(* IEC 61131-3 sources: plcassist-cli/packages/volt-lsp-iec/test-corpus/lenze-mid/Device/Plc Logic/Application/Library Manager/StringUtils, 60 files *)

(* ---- CONSTANTS.gvl ---- *)
VAR_GLOBAL
	NULL : POINTER TO BYTE := 0;
END_VAR

(* ---- GVL_UTF8.gvl ---- *)
VAR_GLOBAL
	TRAILINGBYTESFORUTF8 : ARRAY [0..255] OF BYTE := [0, 0, 0, 0, 0, 0, 0, 0, 0, 0, 0, 0, 0, 0, 0, 0, 0, 0, 0, 0, 0, 0, 0, 0, 0, 0, 0, 0, 0, 0, 0, 0, 0, 0, 0, 0, 0, 0, 0, 0, 0, 0, 0, 0, 0, 0, 0, 0, 0, 0, 0, 0, 0, 0, 0, 0, 0, 0, 0, 0, 0, 0, 0, 0, 0, 0, 0, 0, 0, 0, 0, 0, 0, 0, 0, 0, 0, 0, 0, 0, 0, 0, 0, 0, 0, 0, 0, 0, 0, 0, 0, 0, 0, 0, 0, 0, 0, 0, 0, 0, 0, 0, 0, 0, 0, 0, 0, 0, 0, 0, 0, 0, 0, 0, 0, 0, 0, 0, 0, 0, 0, 0, 0, 0, 0, 0, 0, 0, 0, 0, 0, 0, 0, 0, 0, 0, 0, 0, 0, 0, 0, 0, 0, 0, 0, 0, 0, 0, 0, 0, 0, 0, 0, 0, 0, 0, 0, 0, 0, 0, 0, 0, 0, 0, 0, 0, 0, 0, 0, 0, 0, 0, 0, 0, 0, 0, 0, 0, 0, 0, 0, 0, 0, 0, 0, 0, 0, 0, 0, 0, 0, 0, 1, 1, 1, 1, 1, 1, 1, 1, 1, 1, 1, 1, 1, 1, 1, 1, 1, 1, 1, 1, 1, 1, 1, 1, 1, 1, 1, 1, 1, 1, 1, 1, 2, 2, 2, 2, 2, 2, 2, 2, 2, 2, 2, 2, 2, 2, 2, 2, 3, 3, 3, 3, 3, 3, 3, 3, 4, 4, 4, 4, 5, 5, 5, 5];
	FIRSTBYTEMARK : ARRAY [0..6] OF BYTE := [16#0, 16#0, 16#C0, 16#E0, 16#F0, 16#F8, 16#FC];
	OFFSETSFROMUTF8 : ARRAY [0..5] OF DWORD := [16#0, 16#3080, 16#E2080, 16#3C82080, 16#FA082080, 16#82082080];
	HALFSHIFT : INT := 10;
	HALFBASE : DWORD := 16#10000;
	HALFMASK : DWORD := 16#3FF;
	UNI_REPLACEMENT_CHAR : DWORD := 16#FFFD;
	UNI_MAX_BMP : DWORD := 16#FFFF;
	UNI_MAX_UTF16 : DWORD := 16#10FFFF;
	UNI_MAX_UTF32 : DWORD := 16#7FFFFFFF;
	UNI_MAX_LEGAL_UTF32 : DWORD := 16#10FFFF;
	BYTEMASK : DWORD := 16#BF;
	BYTEMARK : DWORD := 16#80;
	UNI_SUR_HIGH_START : DWORD := 16#D800;
	UNI_SUR_HIGH_END : DWORD := 16#DBFF;
	UNI_SUR_LOW_START : DWORD := 16#DC00;
	UNI_SUR_LOW_END : DWORD := 16#DFFF;
	ERR_SOURCE_EXHAUSTED : UDINT := 16#40A0;
	ERR_TARGET_EXHAUSTED : UDINT := 16#40A1;
	ERR_SOURCE_ILLEGAL : UDINT := 16#40A2;
END_VAR

(* ---- PLACEHOLDERCONSTANTS.gvl ---- *)
VAR_GLOBAL
	DFMT_FIRST_PLACEHOLDER : EDateTimePlaceholder := EDateTimePlaceholder.DFMT_5_DIGIT_DAY;
	DFMT_LAST_PLACEHOLDER : EDateTimePlaceholder := EDateTimePlaceholder.DFMT_1_DIGIT_YEAR;
	TFMT_FIRST_PLACEHOLDER : EDateTimePlaceholder := EDateTimePlaceholder.TFMT_2_DIGIT_HOUR_24_HOUR_CLOCK;
	TFMT_LAST_PLACEHOLDER : EDateTimePlaceholder := EDateTimePlaceholder.TFMT_1_DIGIT_ZONE_DESIGNATOR;
END_VAR

(* ---- STRINGUTILSVERSIONCONSTANTS.gvl ---- *)
VAR_GLOBAL
	_STRINGUTILS_VERSION_LARGEROREQUAL_3_5_3_40_ : INT := 0;
END_VAR

(* ---- ICHARBUFFERSTRING.itf ---- *)
INTERFACE ICHARBUFFERSTRING
END_INTERFACE

METHOD ASWSTRING : CharBufferPtr
END_METHOD

METHOD COPY : DINT
VAR_INPUT
	CBSSOURCE : REFERENCE TO CharBufferString;
END_VAR
END_METHOD

METHOD FROMSTRING : BOOL
VAR_INPUT
	STSTRING : STRING(255);
END_VAR
END_METHOD

METHOD INITCONVERTED : BOOL
VAR_INPUT
	PBUFFER : POINTER TO BYTE;
	UIBUFFERSIZE : UINT;
END_VAR
END_METHOD

(* ---- ILOCALIZEDDATETIMENAMES.itf ---- *)
INTERFACE ILOCALIZEDDATETIMENAMES
END_INTERFACE

METHOD GETDAYLONG : CharBufferPtr
VAR_INPUT
	UIDAYOFWEEK : UINT;
END_VAR
END_METHOD

METHOD GETDAYSHORT : CharBufferPtr
VAR_INPUT
	UIDAYOFWEEK : UINT;
END_VAR
END_METHOD

METHOD GETMONTHLONG : CharBufferPtr
VAR_INPUT
	UIMONTH : UINT;
END_VAR
END_METHOD

METHOD GETMONTHSHORT : CharBufferPtr
VAR_INPUT
	UIMONTH : UINT;
END_VAR
END_METHOD

(* ---- _PRINTF.fun ---- *)
FUNCTION _PRINTF : BOOL
VAR_INPUT
	CBPRESULT : CharBufferPtr;
	UIRESULTCAPACITY : UINT;
	STRINGTYPE : __SYSTEM.TYPE_CLASS;
	CBPFORMAT : CharBufferPtr;
	PVALUE : POINTER TO BYTE;
	TYPECLASS : __SYSTEM.TYPE_CLASS;
END_VAR
END_FUNCTION

(* ---- ANALYZEPLACEHOLDERS.fun ---- *)
FUNCTION ANALYZEPLACEHOLDERS : EPlaceholderAnalyzationState
VAR_INPUT
	RCBSMESSAGE : REFERENCE TO CharBufferString;
	PAPLACEHOLDERS : POINTER TO ARRAY [0..0] OF PlaceholderDescription;
	ICOUNTPLACEHOLDERTOCHECK : INT;
	PAPLACEHOLDEROCCURRENCE : POINTER TO ARRAY [0..0] OF DateTimePlaceholderOccurrence;
	SIMAXCOUNTPLACEHOLDERS : SINT;
END_VAR
VAR_OUTPUT
	SICOUNTPLACEHOLDERS : SINT;
END_VAR
END_FUNCTION

(* ---- ANALYZEPLACEHOLDERSDATETIME.fun ---- *)
FUNCTION ANALYZEPLACEHOLDERSDATETIME : EPlaceholderAnalyzationState
VAR_INPUT
	RCBSMESSAGE : REFERENCE TO CharBufferString;
	PAPLACEHOLDERS : POINTER TO ARRAY [0..0] OF PlaceholderDescription;
	ICOUNTPLACEHOLDERTOCHECK : INT;
	PAPLACEHOLDEROCCURRENCE : POINTER TO ARRAY [0..0] OF DateTimePlaceholderOccurrence;
	SIMAXCOUNTPLACEHOLDERS : SINT;
END_VAR
VAR_OUTPUT
	SICOUNTPLACEHOLDERS : SINT;
END_VAR
END_FUNCTION

(* ---- CHARACTERATEQUALS.fun ---- *)
FUNCTION CHARACTERATEQUALS : BOOL
VAR_INPUT
	CBSSOURCE : REFERENCE TO CharBufferString;
	IPOSITION : INT;
	STCHAR : STRING(1);
END_VAR
END_FUNCTION

(* ---- CHARTOUPPER.fun ---- *)
FUNCTION CHARTOUPPER : BYTE
VAR_INPUT
	BYCHAR : BYTE;
END_VAR
END_FUNCTION

(* ---- CONVERTUTF16TOUTF8.fun ---- *)
FUNCTION CONVERTUTF16TOUTF8 : UDINT
VAR_INPUT
	SOURCESTART : POINTER TO WORD;
	TARGETSTART : POINTER TO BYTE;
	DWTARGETBUFFERSIZE : DWORD;
	BSTRICTCONVERSION : BOOL;
END_VAR
END_FUNCTION

(* ---- CONVERTUTF8TOUTF16.fun ---- *)
FUNCTION CONVERTUTF8TOUTF16 : UDINT
VAR_INPUT
	SOURCESTART : POINTER TO BYTE;
	TARGETSTART : POINTER TO WORD;
	DWTARGETBUFFERSIZE : DWORD;
	BSTRICTCONVERSION : BOOL;
END_VAR
END_FUNCTION

(* ---- HELPISSAMEIGNORECASE.fun ---- *)
FUNCTION HELPISSAMEIGNORECASE : BOOL
VAR_INPUT
	BY1 : BYTE;
	BY2 : BYTE;
END_VAR
END_FUNCTION

(* ---- HELPSTRCMPENDA.fun ---- *)
FUNCTION HELPSTRCMPENDA : BOOL
VAR_INPUT
	PCOMPLETETEXT : CharBufferPtr;
	PSUBTEXT : CharBufferPtr;
	XIGNORECASE : BOOL;
END_VAR
END_FUNCTION

(* ---- HELPSTRCMPSTARTA.fun ---- *)
FUNCTION HELPSTRCMPSTARTA : BOOL
VAR_INPUT
	PCOMPLETETEXT : CharBufferPtr;
	PSUBTEXT : CharBufferPtr;
	XIGNORECASE : BOOL;
END_VAR
END_FUNCTION

(* ---- HELPTRIM.fun ---- *)
FUNCTION HELPTRIM : POINTER TO BYTE
VAR_INPUT
	PTEXT : CharBufferPtr;
	XTRIMLEFT : BOOL;
END_VAR
END_FUNCTION

(* ---- HELPTRIMW.fun ---- *)
FUNCTION HELPTRIMW : POINTER TO WORD
VAR_INPUT
	PTEXT : CharBufferPtr;
	XTRIMLEFT : BOOL;
END_VAR
END_FUNCTION

(* ---- ISLEGALUTF8.fun ---- *)
FUNCTION ISLEGALUTF8 : BOOL
VAR_INPUT
	SOURCE : POINTER TO BYTE;
	LENGTH : INT;
END_VAR
END_FUNCTION

(* ---- ISSPACECHARACTER.fun ---- *)
FUNCTION ISSPACECHARACTER : BOOL
VAR_INPUT
	WCHARACTER : WORD;
END_VAR
END_FUNCTION

(* ---- STRCASECMPA.fun ---- *)
FUNCTION STRCASECMPA : INT
VAR_INPUT
	PBYTE1 : POINTER TO BYTE;
	PBYTE2 : POINTER TO BYTE;
END_VAR
END_FUNCTION

(* ---- STRCASECMPENDA.fun ---- *)
FUNCTION STRCASECMPENDA : INT
VAR_INPUT
	PSTRING : CharBufferPtr;
	PSUFFIX : CharBufferPtr;
END_VAR
END_FUNCTION

(* ---- STRCASECMPSTARTA.fun ---- *)
FUNCTION STRCASECMPSTARTA : INT
VAR_INPUT
	PSTRING : CharBufferPtr;
	PPREFIX : CharBufferPtr;
END_VAR
END_FUNCTION

(* ---- STRCASECMPW.fun ---- *)
FUNCTION STRCASECMPW : INT
VAR_INPUT
	PWD1 : POINTER TO WORD;
	PWD2 : POINTER TO WORD;
END_VAR
END_FUNCTION

(* ---- STRCASEFINDA.fun ---- *)
FUNCTION STRCASEFINDA : INT
VAR_INPUT
	PST1 : POINTER TO STRING(255);
	PST2 : POINTER TO STRING(255);
	UISEARCHSTART : UINT;
END_VAR
END_FUNCTION

(* ---- STRCASEFINDW.fun ---- *)
FUNCTION STRCASEFINDW : INT
VAR_INPUT
	PST1 : POINTER TO WSTRING(255);
	PST2 : POINTER TO WSTRING(255);
	UISEARCHSTART : UINT;
END_VAR
END_FUNCTION

(* ---- STRCMP.fun ---- *)
FUNCTION STRCMP : DINT
VAR_INPUT
	CBSSTRING1 : REFERENCE TO CharBufferString;
	CBSSTRING2 : REFERENCE TO CharBufferString;
END_VAR
END_FUNCTION

(* ---- STRCMPA.fun ---- *)
FUNCTION STRCMPA : INT
VAR_INPUT
	PBY1 : POINTER TO BYTE;
	PBY2 : POINTER TO BYTE;
END_VAR
END_FUNCTION

(* ---- STRCMPENDA.fun ---- *)
FUNCTION STRCMPENDA : INT
VAR_INPUT
	PSTRING : CharBufferPtr;
	PSUFFIX : CharBufferPtr;
END_VAR
END_FUNCTION

(* ---- STRCMPSTARTA.fun ---- *)
FUNCTION STRCMPSTARTA : INT
VAR_INPUT
	PSTRING : CharBufferPtr;
	PPREFIX : CharBufferPtr;
END_VAR
END_FUNCTION

(* ---- STRCMPW.fun ---- *)
FUNCTION STRCMPW : INT
VAR_INPUT
	PWD1 : POINTER TO WORD;
	PWD2 : POINTER TO WORD;
END_VAR
END_FUNCTION

(* ---- STRCONCATA.fun ---- *)
FUNCTION STRCONCATA : BOOL
VAR_INPUT
	PSTFROM : CharBufferPtr;
	PSTTO : CharBufferPtr;
	IBUFFERSIZE : INT;
END_VAR
END_FUNCTION

(* ---- STRCONCATW.fun ---- *)
FUNCTION STRCONCATW : BOOL
VAR_INPUT
	PSTFROM : CharBufferPtr;
	PSTTO : CharBufferPtr;
	IBUFFERSIZE : INT;
END_VAR
END_FUNCTION

(* ---- STRCPY.fun ---- *)
FUNCTION STRCPY : DINT
VAR_INPUT
	CBSTARGET : REFERENCE TO CharBufferString;
	CBSSOURCE : REFERENCE TO CharBufferString;
END_VAR
END_FUNCTION

(* ---- STRCPYA.fun ---- *)
FUNCTION STRCPYA : DINT
VAR_INPUT
	PBUFFER : CharBufferPtr;
	IBUFFERSIZE : DINT;
	PSTR : CharBufferPtr;
END_VAR
END_FUNCTION

(* ---- STRCPYFROM.fun ---- *)
FUNCTION STRCPYFROM : DINT
VAR_INPUT
	RCBSTARGET : REFERENCE TO CharBufferString;
	RCBSSOURCE : REFERENCE TO CharBufferString;
	DISOURCEOFFSET : DINT;
	DITARGETOFFSET : DINT;
	DICOUNTCHARACTERS : DINT;
END_VAR
END_FUNCTION

(* ---- STRCPYW.fun ---- *)
FUNCTION STRCPYW : DINT
VAR_INPUT
	PBUFFER : CharBufferPtr;
	IBUFFERSIZE : DINT;
	PSTR : CharBufferPtr;
END_VAR
END_FUNCTION

(* ---- STRFIND.fun ---- *)
FUNCTION STRFIND : INT
VAR_INPUT
	CBSSOURCE : REFERENCE TO CharBufferString;
	CBSTOSEARCHFOR : REFERENCE TO CharBufferString;
END_VAR
END_FUNCTION

(* ---- STRFINDA.fun ---- *)
FUNCTION STRFINDA : INT
VAR_INPUT
	PST1 : POINTER TO STRING(255);
	PST2 : POINTER TO STRING(255);
	UISEARCHSTART : UINT;
END_VAR
END_FUNCTION

(* ---- STRFINDFROM.fun ---- *)
FUNCTION STRFINDFROM : INT
VAR_INPUT
	CBSSOURCE : REFERENCE TO CharBufferString;
	CBSTOSEARCHFOR : REFERENCE TO CharBufferString;
	ISEARCHSTART : UINT;
END_VAR
END_FUNCTION

(* ---- STRFINDW.fun ---- *)
FUNCTION STRFINDW : INT
VAR_INPUT
	PST1 : POINTER TO WSTRING(255);
	PST2 : POINTER TO WSTRING(255);
	UISEARCHSTART : UINT;
END_VAR
END_FUNCTION

(* ---- STRINGTOCHARBUFFERPTR.fun ---- *)
FUNCTION STRINGTOCHARBUFFERPTR : BOOL
VAR_INPUT
	STSTRING : STRING(255);
	CBSRESULT : REFERENCE TO CharBufferString;
END_VAR
END_FUNCTION

(* ---- STRISNULLOREMPTYA.fun ---- *)
FUNCTION STRISNULLOREMPTYA : BOOL
VAR_INPUT
	PSTDATA : CharBufferPtr;
END_VAR
END_FUNCTION

(* ---- STRISNULLOREMPTYW.fun ---- *)
FUNCTION STRISNULLOREMPTYW : BOOL
VAR_INPUT
	PSTDATA : CharBufferPtr;
END_VAR
END_FUNCTION

(* ---- STRLEN.fun ---- *)
FUNCTION STRLEN : DINT
VAR_INPUT
	CBSSOURCE : REFERENCE TO CharBufferString;
END_VAR
END_FUNCTION

(* ---- STRLENA.fun ---- *)
FUNCTION STRLENA : DINT
VAR_INPUT
	PSTDATA : CharBufferPtr;
END_VAR
END_FUNCTION

(* ---- STRLENW.fun ---- *)
FUNCTION STRLENW : DINT
VAR_INPUT
	PSTDATA : CharBufferPtr;
END_VAR
END_FUNCTION

(* ---- STRPADLEFTA.fun ---- *)
FUNCTION STRPADLEFTA : BOOL
VAR_INPUT
	BYPADCHAR : BYTE;
	PSTFROM : CharBufferPtr;
	PSTTO : CharBufferPtr;
	DIBUFFERSIZE : DINT;
END_VAR
END_FUNCTION

(* ---- STRPADLEFTW.fun ---- *)
FUNCTION STRPADLEFTW : BOOL
VAR_INPUT
	WPADCHAR : WORD;
	PSTFROM : CharBufferPtr;
	PSTTO : CharBufferPtr;
	DIBUFFERSIZE : DINT;
END_VAR
END_FUNCTION

(* ---- STRPADRIGHTA.fun ---- *)
FUNCTION STRPADRIGHTA : BOOL
VAR_INPUT
	BYPADCHAR : BYTE;
	PSTFROM : CharBufferPtr;
	PSTTO : CharBufferPtr;
	DIBUFFERSIZE : DINT;
END_VAR
END_FUNCTION

(* ---- STRPADRIGHTW.fun ---- *)
FUNCTION STRPADRIGHTW : BOOL
VAR_INPUT
	WPADCHAR : WORD;
	PSTFROM : CharBufferPtr;
	PSTTO : CharBufferPtr;
	DIBUFFERSIZE : DINT;
END_VAR
END_FUNCTION

(* ---- STRTRIMW.fun ---- *)
FUNCTION STRTRIMW : BOOL
VAR_INPUT
	PSTRING : CharBufferPtr;
END_VAR
END_FUNCTION

(* ---- STUSPRINTF.fun ---- *)
FUNCTION STUSPRINTF : INT
VAR_INPUT
	PSTFORMAT : POINTER TO STRING;
	PVARADR : POINTER TO DWORD;
	UDIVARTYPE : __SYSTEM.TYPE_CLASS;
	PBUFFER : POINTER TO BYTE;
	DWBUFFERSIZE : UDINT;
END_VAR
END_FUNCTION

(* ---- STUSPRINTFW.fun ---- *)
FUNCTION STUSPRINTFW : INT
VAR_INPUT
	WSTFORMAT : POINTER TO WSTRING;
	PVARADR : POINTER TO DWORD;
	UDIVARTYPE : __SYSTEM.TYPE_CLASS;
	PBUFFER : POINTER TO BYTE;
	DWBUFFERSIZE : UDINT;
END_VAR
END_FUNCTION

(* ---- WCHARTOUPPER.fun ---- *)
FUNCTION WCHARTOUPPER : WORD
VAR_INPUT
	WDCHAR : WORD;
END_VAR
END_FUNCTION

(* ---- ABSTRACTFORMATTER.fb ---- *)
FUNCTION_BLOCK ABSTRACTFORMATTER
VAR
	M_APLACEHOLDEROCCURRENCE : ARRAY [0..(COUNT_PLACEHOLDERS_IN_FORMAT_STRING - 1)] OF DateTimePlaceholderOccurrence;
	M_SICOUNTPLACEHOLDERS : SINT := -1;
	M_EPLACEHOLDERANALYZATIONSTATE : EPlaceholderAnalyzationState;
	M_SFORMATSTRING : STRING(50);
	M_IFORMATSTRINGLENGTH : INT;
	COUNT_PLACEHOLDERS_IN_FORMAT_STRING : INT := 10;
	COUNT_PLACEHOLDERS_IN_DATETIMEFORMAT_STRING : INT := 20;
	MAX_FORMAT_STRING_LENGTH : SINT := 50;
END_VAR
END_FUNCTION_BLOCK

(* ---- CHARBUFFERSTRING.fb ---- *)
FUNCTION_BLOCK CHARBUFFERSTRING
VAR_INPUT
	M_UIBUFFERSIZE : UINT;
	M_CBPBUFFER : CharBufferPtr;
	M_TYPE : __SYSTEM.TYPE_CLASS;
	M_ASSTRING : POINTER TO STRING(255);
	M_ASWSTRING : POINTER TO WSTRING(255);
	M_BALLOCATED : BOOL;
END_VAR
VAR
	CAPACITY : UINT;
	CHARACTERS : CharBufferPtr;
	LENGTH : DINT;
	STRINGTYPE : __SYSTEM.TYPE_CLASS;
END_VAR
END_FUNCTION_BLOCK

METHOD ASWSTRING : CharBufferPtr
END_METHOD

METHOD CHARAT : BYTE
VAR_INPUT
	IPOSITION : INT;
END_VAR
END_METHOD

METHOD CHARATEQUALS : BOOL
VAR_INPUT
	IPOSITION : INT;
	STCHAR : STRING(1);
END_VAR
END_METHOD

METHOD COPY : DINT
VAR_INPUT
	CBSSOURCE : REFERENCE TO CharBufferString;
END_VAR
END_METHOD

METHOD COPYFROM
VAR_INPUT
	RCBSSOURCE : REFERENCE TO CharBufferString;
	DISOURCEOFFSET : DINT;
	DITARGETOFFSET : DINT;
	DICOUNTCHARACTERS : DINT;
END_VAR
END_METHOD

METHOD COPYFROM2 : DINT
VAR_INPUT
	RSSOURCE : REFERENCE TO STRING(255);
	DITARGETOFFSET : DINT;
END_VAR
END_METHOD

METHOD DELETE : DINT
VAR_INPUT
	ILENGTH : INT;
	IPOSITION : INT;
END_VAR
END_METHOD

METHOD FB_EXIT : BOOL
VAR_INPUT
	BINCOPYCODE : BOOL;
END_VAR
END_METHOD

METHOD FB_INIT : BOOL
VAR_INPUT
	BINITRETAINS : BOOL;
	BINCOPYCODE : BOOL;
	UIBUFFERSIZE : UINT;
	STRINGTYPE : __SYSTEM.TYPE_CLASS;
END_VAR
END_METHOD

METHOD FIND : INT
VAR_INPUT
	CBSTOSEARCHFOR : REFERENCE TO CharBufferString;
END_VAR
END_METHOD

METHOD FINDFROM : INT
VAR_INPUT
	CBSTOSEARCHFOR : REFERENCE TO CharBufferString;
	ISEARCHSTART : UINT;
END_VAR
END_METHOD

METHOD FROMSTRING : BOOL
VAR_INPUT
	STSTRING : STRING(255);
END_VAR
END_METHOD

METHOD INIT : BOOL
VAR_INPUT
	PBUFFER : POINTER TO BYTE;
	UIBUFFERSIZE : UINT;
	STRINGTYPE : __SYSTEM.TYPE_CLASS;
END_VAR
END_METHOD

METHOD INITCONVERTED : BOOL
VAR_INPUT
	PBUFFER : POINTER TO BYTE;
	UIBUFFERSIZE : UINT;
END_VAR
END_METHOD

METHOD INITIALIZE : BOOL
VAR_INPUT
	CBPSOURCE : CharBufferPtr;
	STRINGTYPE : __SYSTEM.TYPE_CLASS;
END_VAR
END_METHOD

METHOD INSERT
VAR_INPUT
	CBSINSERT : REFERENCE TO CharBufferString;
	IPOSITION : INT;
END_VAR
END_METHOD

METHOD MID
VAR_INPUT
	ILENGTH : INT;
	IPOSITION : INT;
	CBSRESULT : REFERENCE TO CharBufferString;
END_VAR
END_METHOD

METHOD PLACEHOLDEREQUALS : BOOL
VAR_INPUT
	STVALUE : STRING;
	WSTVALUE : WSTRING;
END_VAR
END_METHOD

METHOD REPLACE
VAR_INPUT
	CBSREPLACEWITH : REFERENCE TO CharBufferString;
	ILENGTHTOREPLACE : INT;
	IPOSITION : INT;
END_VAR
END_METHOD

(* ---- DATEFORMATTER.fb ---- *)
FUNCTION_BLOCK DATEFORMATTER EXTENDS AbstractFormatter
VAR
	M_CBSPLACEHOLDER2DIGITDAY : CharBufferString;
	M_CBSPLACEHOLDER1DIGITDAY : CharBufferString;
	M_CBSPLACEHOLDER2DIGITMONTH : CharBufferString;
	M_CBSPLACEHOLDER1DIGITMONTH : CharBufferString;
	M_CBSPLACEHOLDER4DIGITYEAR : CharBufferString;
	M_CBSPLACEHOLDER2DIGITYEAR : CharBufferString;
	M_CBSPLACEHOLDER1DIGITYEAR : CharBufferString;
END_VAR
END_FUNCTION_BLOCK

METHOD FB_EXIT : BOOL
VAR_INPUT
	BINCOPYCODE : BOOL;
END_VAR
END_METHOD

METHOD FB_INIT : BOOL
VAR_INPUT
	BINITRETAINS : BOOL;
	BINCOPYCODE : BOOL;
END_VAR
END_METHOD

METHOD FORMAT : STRING
VAR_INPUT
	PDATE : SYSTIMEDATE;
END_VAR
END_METHOD

METHOD SETFORMATSTRING
VAR_INPUT
	SFORMATSTRING : STRING(MAX_FORMAT_STRING_LENGTH);
END_VAR
END_METHOD

(* ---- DATETIMEFORMATTER.fb ---- *)
FUNCTION_BLOCK DATETIMEFORMATTER EXTENDS AbstractFormatter
VAR
	M_APLACEHOLDEROCCURRENCEDATETIME : ARRAY [0..(COUNT_PLACEHOLDERS_IN_DATETIMEFORMAT_STRING - 1)] OF DateTimePlaceholderOccurrence;
	M_CBSPLACEHOLDER5DIGITDAY : CharBufferString;
	M_CBSPLACEHOLDER4DIGITDAY : CharBufferString;
	M_CBSPLACEHOLDER3DIGITDAY : CharBufferString;
	M_CBSPLACEHOLDER2DIGITDAY : CharBufferString;
	M_CBSPLACEHOLDER1DIGITDAY : CharBufferString;
	M_CBSPLACEHOLDER3DIGITDAYOFYEAR : CharBufferString;
	M_CBSPLACEHOLDER4DIGITMONTH : CharBufferString;
	M_CBSPLACEHOLDER3DIGITMONTH : CharBufferString;
	M_CBSPLACEHOLDER2DIGITMONTH : CharBufferString;
	M_CBSPLACEHOLDER1DIGITMONTH : CharBufferString;
	M_CBSPLACEHOLDER4DIGITYEAR : CharBufferString;
	M_CBSPLACEHOLDER2DIGITYEAR : CharBufferString;
	M_CBSPLACEHOLDER1DIGITYEAR : CharBufferString;
	M_CBSPLACEHOLDER2DIGITHOUR24HOURCLOCK : CharBufferString;
	M_CBSPLACEHOLDER1DIGITHOUR24HOURCLOCK : CharBufferString;
	M_CBSPLACEHOLDER2DIGITHOUR12HOURCLOCK : CharBufferString;
	M_CBSPLACEHOLDER1DIGITHOUR12HOURCLOCK : CharBufferString;
	M_CBSPLACEHOLDER2DIGITMINUTE : CharBufferString;
	M_CBSPLACEHOLDER1DIGITMINUTE : CharBufferString;
	M_CBSPLACEHOLDER2DIGITSECOND : CharBufferString;
	M_CBSPLACEHOLDER1DIGITSECOND : CharBufferString;
	M_CBSPLACEHOLDER3DIGITMILLISECOND : CharBufferString;
	M_CBSPLACEHOLDER3DIGITMICROSECOND : CharBufferString;
	M_CBSPLACEHOLDER3DIGITNANOSECOND : CharBufferString;
	M_CBSPLACEHOLDER2DIGITAMPMDESIGNATOR : CharBufferString;
	M_CBSPLACEHOLDER1DIGITAMPMDESIGNATOR : CharBufferString;
	M_CBSPLACEHOLDER1DIGITZONEDESIGNATOR : CharBufferString;
	M_OPTLOCALIZER : ILocalizedDateTimeNames;
	M_IUTCOFFSET : INT;
END_VAR
END_FUNCTION_BLOCK

METHOD FB_EXIT : BOOL
VAR_INPUT
	BINCOPYCODE : BOOL;
END_VAR
END_METHOD

METHOD FB_INIT : BOOL
VAR_INPUT
	BINITRETAINS : BOOL;
	BINCOPYCODE : BOOL;
END_VAR
END_METHOD

METHOD FORMAT : WSTRING
VAR_INPUT
	PDATE : SYSTIMEDATE;
	UIMICROSECONDS : UINT;
	UINANOSECONDS : UINT;
	DATATYPE : __SYSTEM.TYPE_CLASS := __SYSTEM.TYPE_CLASS.TYPE_NONE;
END_VAR
END_METHOD

METHOD FORMATSINGLEDIGIT : WSTRING
VAR_INPUT
	PDATE : SYSTIMEDATE;
	UIMICROSECONDS : UINT;
	UINANOSECONDS : UINT;
	DATATYPE : __SYSTEM.TYPE_CLASS := __SYSTEM.TYPE_CLASS.TYPE_NONE;
	SIINDEXOFSINGLEDIGITTORETURN : SINT;
END_VAR
VAR_OUTPUT
	ICOPYSINGLETARGETOFFSET : INT;
END_VAR
END_METHOD

METHOD FORMATWITHUTCOFFSET : WSTRING
VAR_INPUT
	PDATE : SYSTIMEDATE;
	UIMICROSECONDS : UINT;
	UINANOSECONDS : UINT;
	DATATYPE : __SYSTEM.TYPE_CLASS := __SYSTEM.TYPE_CLASS.TYPE_NONE;
	IUTCOFFSET : INT;
END_VAR
END_METHOD

METHOD SETFORMATSTRING
VAR_INPUT
	SFORMATSTRING : STRING(MAX_FORMAT_STRING_LENGTH);
END_VAR
END_METHOD

METHOD SETLOCALIZER
VAR_INPUT
	LOCALIZER : ILocalizedDateTimeNames;
END_VAR
END_METHOD

METHOD GETDAY : WSTRING
VAR_INPUT
	UIDAYOFWEEK : UINT;
	DAYFORMAT : EDateTimePlaceholder;
END_VAR
VAR_IN_OUT
	DILENGTH : DINT;
END_VAR
END_METHOD

METHOD GETMONTH : WSTRING
VAR_INPUT
	UIMONTH : UINT;
	MONTHFORMAT : EDateTimePlaceholder;
END_VAR
VAR_IN_OUT
	DILENGTH : DINT;
END_VAR
END_METHOD

(* ---- TIMEFORMATTER.fb ---- *)
FUNCTION_BLOCK TIMEFORMATTER EXTENDS AbstractFormatter
VAR
	M_CBSPLACEHOLDER2DIGITHOUR24HOURCLOCK : CharBufferString;
	M_CBSPLACEHOLDER1DIGITHOUR24HOURCLOCK : CharBufferString;
	M_CBSPLACEHOLDER2DIGITHOUR12HOURCLOCK : CharBufferString;
	M_CBSPLACEHOLDER1DIGITHOUR12HOURCLOCK : CharBufferString;
	M_CBSPLACEHOLDER2DIGITMINUTE : CharBufferString;
	M_CBSPLACEHOLDER1DIGITMINUTE : CharBufferString;
	M_CBSPLACEHOLDER2DIGITSECOND : CharBufferString;
	M_CBSPLACEHOLDER1DIGITSECOND : CharBufferString;
	M_CBSPLACEHOLDER3DIGITMILLISECOND : CharBufferString;
	M_CBSPLACEHOLDER3DIGITMICROSECOND : CharBufferString;
	M_CBSPLACEHOLDERAMPMDESIGNATOR : CharBufferString;
	M_CBSPLACEHOLDER1DIGITZONEDESIGNATOR : CharBufferString;
END_VAR
END_FUNCTION_BLOCK

METHOD FB_EXIT : BOOL
VAR_INPUT
	BINCOPYCODE : BOOL;
END_VAR
END_METHOD

METHOD FB_INIT : BOOL
VAR_INPUT
	BINITRETAINS : BOOL;
	BINCOPYCODE : BOOL;
END_VAR
END_METHOD

METHOD FORMAT : STRING
VAR_INPUT
	PDATE : SYSTIMEDATE;
	UIMIRCOSECONDS : UINT;
END_VAR
END_METHOD

METHOD FORMATWITHUTCOFFSET : STRING
VAR_INPUT
	PDATE : SYSTIMEDATE;
	UIMIRCOSECONDS : UINT;
	IUTCOFFSET : INT;
END_VAR
END_METHOD

METHOD SETFORMATSTRING
VAR_INPUT
	SFORMATSTRING : STRING(MAX_FORMAT_STRING_LENGTH);
END_VAR
END_METHOD
